Fanuc KAREL source: ka00144.KL

-- PROVISIONAL review KL for V1013-1; original PC SHA256 904954391d082d173cf3ea4f97d9d3371533677b5027ef5598d3815056e34669
-- Incomplete behavior may be omitted. Consult companion uncertainty JSON. Do not deploy.
PROGRAM KA00144
%NOLOCKGROUP
-- UNRESOLVED_DECL SRC type=002017
-- UNRESOLVED_DECL DST type=002017
BEGIN
  -- UNRESOLVED_PC offsets 5-19; opcodes 2E,22,9D,33,B4
  -- UNRESOLVED_PC offsets 24-42; opcodes 22,9D,33,B3,22,9D,33,B4
  -- UNRESOLVED_PC offsets 47-51; opcodes 7F
END KA00144
